{attribute 'qualified_only'}
{attribute 'strict'}
{attribute 'to_string'}
TYPE E_HMIKistlerResult :
(
    NONE := 0,
    PASS := 1,
    FAIL := 2
);
END_TYPE

(* stored: Version 1.1.0.1
   DUT E_HMIKistlerResult: Id {3b73df06-8057-4b20-b1eb-1c4fa9c6670d} *)
